Fanuc KAREL source: KT00711.KL

PROGRAM KT00711
%NOLOCKGROUP
VAR
  B1: BOOLEAN
  B2: BOOLEAN
  OUT: INTEGER
BEGIN
  B1 = TRUE
  B2 = FALSE
  B1 = TRUE
  B2 = FALSE
  OUT = ARRAY_LEN(B1)
END KT00711
